(* IEC 61131-3 sources: codesys-to-astra/cds2astra/tests/corpus/C2A-LIB001/pos/src/POUs/PRG_A, 1 file *)

(* ---- PRG_A.decl.st ---- *)
// Назначение: корпус правила cds2astra (synthetic).
// Автор:      kr0nsch
// Версия:     0.1.0
// Документ:   docs/RULES.md
PROGRAM PRG_A
VAR
    sHex : STRING(8); // строка
END_VAR
